Universal Robots URScript: JointTargets.script

def JointTargets():
  # Global parameters:
  global speed_ms    = 0.250
  global speed_rads  = 0.750
  global accel_mss   = 1.200
  global accel_radss = 1.200
  global blend_radius_m = 0.001
  global ref_frame = p[0,0,0,0,0,0]

  #
  # TO REMOVE HEADER:
  # Go to "Program" -> "Post-Processor Editor"
  # Select "Universal Robots"
  # Set "INCLUDE_HEADER" to "False"
  #
  #--------------------------
  # Add any default subprograms here
  # For example, to drive a gripper as a program call:
  # def Gripper_Open():
  #   ...
  # end
  #
  # Example to drive a spray gun:
  def SprayOn(value):
    # use the value as an output:
    DO_SPRAY = 5
    if value == 0:
      set_standard_digital_out(DO_SPRAY, False)
    else:
      set_standard_digital_out(DO_SPRAY, True)
    end
  end

  # Example to drive an extruder:
  def Extruder(value):
    # use the value as an output:
    if value < 0:
      # stop extruder
    else:
      # start extruder
    end
  end

  # Example to move an external axis
  def MoveAxis(value):
    # use the value as an output:
    DO_AXIS_1 = 1
    DI_AXIS_1 = 1
    if value <= 0:
      set_standard_digital_out(DO_AXIS_1, False)

      # Wait for digital input to change state
      #while (get_standard_digital_in(DI_AXIS_1) != False):
      #  sync()
      #end
    else:
      set_standard_digital_out(DO_AXIS_1, True)

      # Wait for digital input to change state
      #while (get_standard_digital_in(DI_AXIS_1) != True):
      #  sync()
      #end
    end
  end
  #--------------------------


  # Main program:
  # Program generated by VerticalBot Studio for UR5e on 25/10/2026 12:00:00
  # Using nominal kinematics.
  ref_frame = p[0.100000, -0.050000, 0.020000, 0.000000, 0.000000, 0.523599]
  set_tcp(p[0.010000, 0.000000, 0.120000, 0.000000, 0.261799, 0.000000])
  movej([-0.523599, -1.745329, 1.570796, -1.396263, -1.570796, 0.349066],accel_radss,speed_rads,0,0)
  movel([-0.383972, -1.675516, 1.570796, -1.396263, -1.570796, 0.349066],accel_mss,speed_ms,0,0)
  movej([-0.383972, -1.675516, 1.570796, -1.396263, -1.570796, 0.349066],accel_radss,speed_rads,0,0.001)
  movel(pose_trans(ref_frame,p[-0.373291, 0.385355, 0.409557, -3.080591, -0.269517, -0.405567]),accel_mss,speed_ms,0,0.001)
  movel([-0.383972, -1.675516, 1.570796, -1.396263, -1.570796, 0.349066],accel_mss,speed_ms,0,0)
  blend_radius_m = 0.005
  movej([-0.523599, -1.745329, 1.570796, -1.396263, -1.570796, 0.349066],accel_radss,speed_rads,0,0)
  movel([-0.383972, -1.675516, 1.570796, -1.396263, -1.570796, 0.349066],accel_mss,speed_ms,0,0)
  movej([-0.383972, -1.675516, 1.570796, -1.396263, -1.570796, 0.349066],accel_radss,speed_rads,0,0.005)
  movel(pose_trans(ref_frame,p[-0.373291, 0.385355, 0.409557, -3.080591, -0.269517, -0.405567]),accel_mss,speed_ms,0,0.005)
  movel([-0.383972, -1.675516, 1.570796, -1.396263, -1.570796, 0.349066],accel_mss,speed_ms,0,0)
  blend_radius_m = 0.000
  movej([-0.523599, -1.745329, 1.570796, -1.396263, -1.570796, 0.349066],accel_radss,speed_rads,0,0)
  # End of main program
end

JointTargets()
